Fanuc KAREL source: KC00026.KL

PROGRAM KC00026
%NOLOCKGROUP
%ENVIRONMENT UIF
VAR
  I: INTEGER
  J: INTEGER
  K: INTEGER
  R: REAL
  B: BOOLEAN
  S: STRING[80]
  T: STRING[80]
  P: PATH
  Q: PATH
  AI: ARRAY[8] OF INTEGER
  AB: ARRAY[244] OF BYTE
  X: XWORK_T
BEGIN
  ACT_TBL(I,J,X,K,B,I)
END KC00026
